Staubli VAL3: HMI_progEdit.pjx

--- HMI_progEdit.pjx ---
Parameters version=s8.12.2Cs9_BS2561 stackSize=5000 millimeterUnit=true
Program file=_bindPROG.pgx
Program file=_bindTRAJ.pgx
Program file=_btnColor.pgx
Program file=_onStartPROG.pgx
Program file=_onStartTRAJ.pgx
Program file=bind.pgx
Program file=IFedit.pgx
Program file=insertCASE.pgx
Program file=insertFOR.pgx
Program file=insertIF.pgx
Program file=insertSwitch.pgx
Program file=insetProg.pgx
Program file=main.pgx
Program file=onStart.pgx
Program file=refreshlist.pgx
Program file=resfreshPROG.pgx
Program file=resfreshTRAJ.pgx
Program file=start.pgx
Program file=stop.pgx
Program file=unbind.pgx
Data file=HMI_progEdit.dtx
Library alias=rs path=Disk://source/projectSource/robotStatus/robotStatus.pjx
Library alias=prog path=Disk://source/projectSource/program/program.pjx
Library alias=util path=Disk://HMI_cs9/HMI_util/HMI_util.pjx
Library alias=progTemp path=Disk://source/template/progTemp/progTemp.pjx
Library alias=simulate path=Disk://HMI_cs9/simulate/simulate.pjx
Library alias=trajectory path=Disk://source/projectSource/trajectory/trajectory.pjx
Library alias=io path=Disk://source/projectSource/io/io.pjx

--- HMI_progEdit.dtx ---
mdesc mNomSpeed
string sSelProg
bool bBack
public bool bBool[9]
public bool bInsert[16]
num nPageIndex
num nPageNum
public num nLstValue
string sLstValue
string sList
bool bToSave
string sPageNum
string sPageIndex
public bool bTRAJ[7]
string sPgIndexTRAJ
string sPageTRAJ
num nPgIndexTRAJ
num nPgNumTRAJ
string sTRAJList
string sInsertItem
string sPgIndexPROG
string sPagePROG
num nPgIndexPROG
num nPgNumPROG
string sPROGList
string sIFType[3]
public num nIFValue[3]
string sIFIndex[3]
string sANDOR1
string sANDOR2
bool bIFConfirm
bool bIFCancel
string sLastANDOR2
string sLastANDOR1
bool bSwitchOK
bool bSwitchCancel
string sIOList
string sSwitchValue
num nCaseValue
num nFORValue
string sForValue
bool bSelProg
bool bSelTraj
bool bBindTRAJ
bool bBindProg
num nSelType

--- main.pgx ---
public program main(string x_sSelProg)
  local bool l_bExit
  local bool l_bRefresh
  local num l_nIndex
begin
  //x_sSelProg-选中的prog
  do
    if util:sPage!="editProg"
      util:sPage="editProg"
      sSelProg= x_sSelProg
      call onStart()
      call bind()
      userPage(util:sPage)
      delay(0.5)
      l_bRefresh=true
    endIf

    if bBool[1]
      bBool[1]=false
      call simulate:simulatePROG(sSelProg)
    elseIf bBool[2]
      bBool[2]=false
      call prog:deleteProgItem(sSelProg,sLstValue,bToSave)
      l_bRefresh=true
    elseIf bBool[3]
      bBool[3]=false

    elseIf bBool[4]
      bBool[4]=false
      progTemp:libSave()
      delay(0.1)
      popUpMsg("数据已保存")
    elseIf bBool[5]
      bBool[5]=false
      nPageIndex=0
      l_bRefresh=true
    elseIf bBool[6]
      bBool[6]=false
      if nPageIndex>0
        nPageIndex=nPageIndex-1
      endIf
      l_bRefresh=true
    elseIf bBool[7]
      bBool[7]=false
      if nPageIndex<nPageNum-1
        nPageIndex=nPageIndex+1
      endIf
      l_bRefresh=true
    elseIf bBool[8]
      bBool[8]=false
      nPageIndex=nPageNum-1
      l_bRefresh=true
    elseIf bInsert[0]
      bInsert[0]=false
      call unbind()
      call prog:getProgItemIndex(sSelProg,sLstValue,l_nIndex)
      //call insetTRAJ(l_nIndex)
      l_bRefresh=true
    elseIf bInsert[1]
      bInsert[1]=false
      call unbind()
      call prog:getProgItemIndex(sSelProg,sLstValue,l_nIndex)
      call insetProg(l_nIndex,bToSave)
      l_bRefresh=true
    elseIf bInsert[2]
      bInsert[2]=false
      call insertIF()
      l_bRefresh=true
    elseIf bInsert[3]
      bInsert[3]=false
      call prog:getProgItemIndex(sSelProg,sLstValue,l_nIndex)
      call prog:insertENDIF(sSelProg,l_nIndex,bToSave)
      l_bRefresh=true
    elseIf bInsert[4]
      bInsert[4]=false
      call insertSwitch()
      l_bRefresh=true
    elseIf bInsert[5]
      bInsert[5]=false
      call prog:getProgItemIndex(sSelProg,sLstValue,l_nIndex)
      call insertCASE(l_nIndex)
      l_bRefresh=true
    elseIf bInsert[6]
      bInsert[6]=false
      call prog:getProgItemIndex(sSelProg,sLstValue,l_nIndex)
      call prog:insertENDSwitch(sSelProg,l_nIndex,bToSave)
      l_bRefresh=true
    elseIf bInsert[7]
      bInsert[7]=false
      call prog:getProgItemIndex(sSelProg,sLstValue,l_nIndex)
      call insertFOR(l_nIndex)
      l_bRefresh=true
    elseIf bBack
      bBack=false
      //call prog:onSave(bToSave)
      l_bExit=true
    endIf

    if l_bRefresh
      l_bRefresh=false
      call refreshlist()

    endIf



    delay(0)
  until l_bExit==true
  if bToSave
    call prog:onSave(bToSave)
  endIf
end

--- start.pgx ---
program start()
begin
end

--- _bindPROG.pgx ---
program _bindPROG(string x_sHtml)
  local num l_i
  local string l_sbtn
begin
  for l_i = 1 to 6
    l_sbtn="btn"+toString("",l_i)
    userPageBindClick(x_sHtml,l_sbtn,bInsert[l_i],true)
  endFor

  userPageBind(x_sHtml,"lbl1","innerHTML",sPgIndexPROG,1,"r")
  userPageBind(x_sHtml,"lbl2","innerHTML",sPagePROG,1,"r")

  userPageBindClick(x_sHtml,"btn7",bSelProg,true)
  userPageBindClick(x_sHtml,"btn8",bSelTraj,true)
  userPageBind(x_sHtml,"lst1","value",sInsertItem,1,"rw")

end

--- _bindTRAJ.pgx ---
program _bindTRAJ()
  local num l_i
  local string l_sbtn
begin
  for l_i = 1 to 6
    l_sbtn="btn"+toString("",l_i)
    userPageBindClick("insertTRAJ",l_sbtn,bInsert[l_i],true)
  endFor

  userPageBind("insertTRAJ","lbl1","innerHTML",sPgIndexTRAJ,1,"r")
  userPageBind("insertTRAJ","lbl2","innerHTML",sPageTRAJ,1,"r")


  userPageBind("insertTRAJ","lst1","value",sInsertItem,1,"rw")
end

--- _btnColor.pgx ---
public program _btnColor(num x_nSelType, string x_sHtml)
begin
  switch x_nSelType
    case 1
      userPageSet(x_sHtml,"btn7","style.backgroundColor","#7CB5FF")
      userPageSet(x_sHtml,"btn7","style.color","#FFFFFF")
      userPageSet(x_sHtml,"btn8","style.backgroundColor","#FFFFFF")
      userPageSet(x_sHtml,"btn8","style.color","#838A8F")
    break
    case 2
      userPageSet(x_sHtml,"btn8","style.backgroundColor","#7CB5FF")
      userPageSet(x_sHtml,"btn8","style.color","#FFFFFF")
      userPageSet(x_sHtml,"btn7","style.backgroundColor","#FFFFFF")
      userPageSet(x_sHtml,"btn7","style.color","#838A8F")
    break
  endSwitch

end

--- _onStartPROG.pgx ---
public program _onStartPROG(string x_sHtml)
begin
  nPgIndexPROG=0
  nPgNumPROG=0
  sPagePROG=""
  sPgIndexPROG=""
  bSelProg=true
  bSelTraj=false
  if bSelProg
    call resfreshPROG(x_sHtml)
  elseIf bSelTraj
    call resfreshTRAJ(x_sHtml)
  endIf
end

--- _onStartTRAJ.pgx ---
public program _onStartTRAJ()
begin
  nPgIndexTRAJ=0
  nPgNumTRAJ=0
  sPageTRAJ=""
  sPgIndexTRAJ=""
//  call resfreshTRAJ()
end

--- bind.pgx ---
program bind()
  local string l_sbtn
  local num l_i
begin
  //button
  userPageBindClick("editProg","btnback",bBack,true)
  for l_i = 1 to 8
    l_sbtn="btn"+toString("",l_i)
    userPageBindClick("editProg",l_sbtn,bBool[l_i],true)
  endFor

  for l_i = 0 to 8
    l_sbtn="btn1"+toString("",l_i)
    userPageBindClick("editProg",l_sbtn,bInsert[l_i],true)
  endFor

  //lbl
  userPageBind("editProg","lbl1","innerHTML",sSelProg,1,"r")
  userPageBind("editProg","lbleditindex","innerHTML",sPageIndex,1,"r")
  userPageBind("editProg","lbleditpage","innerHTML",sPageNum,1,"r")

  //lst
  userPageBind("editProg","lst1","options",sList,size(sList),"r")
  userPageBind("editProg","lst1","value",sLstValue,1,"rw")

end

--- IFedit.pgx ---
program IFedit(num x_nIndex)
begin
  call prog:editIF(sSelProg,x_nIndex,sIFType,sIFIndex,nIFValue,sANDOR1,sANDOR2,bToSave)
end

--- insertCASE.pgx ---
public program insertCASE(num x_nProgIndex)
  local bool l_bExit
  local bool l_bRefreh
  local num l_nProgIndex
  local num l_i
  local bool l_bRefresh
begin
  do
    if util:sPage!="insertCASE"
      util:sPage="insertCASE"
      call _onStartPROG(util:sPage)
      call _bindPROG(util:sPage)
      userPageBind("insertCASE","nmb1","value",nCaseValue,1,"rw")
      if size(sIOList)!=(size(io:aInItem)+1)
        resize(sIOList,1,size(io:aInItem)+1)
      endIf
      for l_i = 1 to size(sIOList)-1
        sIOList[l_i-1]=toString("",l_i-1)+","+io:aInItem[l_i-1].sComment
      endFor
      sIOList[0]=""
      userPage(util:sPage)
      delay(0.5)
    endIf

    //btn
    if bSelProg
      bSelProg=false
      nSelType=1
      l_bRefresh=true
      nPgIndexPROG=0
    elseIf bSelTraj
      bSelTraj=false
      nSelType=2
      l_bRefresh=true
      nPgIndexPROG=0
    endIf

    //refresh
    if l_bRefresh
      l_bRefresh=false
      call _btnColor(nSelType,util:sPage)
      switch nSelType
        case 1
          call resfreshPROG(util:sPage)
        break
        case 2
          nPgIndexTRAJ=0
          call resfreshTRAJ(util:sPage)
        break
      endSwitch
    endIf

    if bInsert[1]
      bInsert[1]=false

      call prog:insertCASE(sSelProg,x_nProgIndex,sInsertItem,bToSave,nCaseValue,nSelType)

      l_bExit=true
    elseIf bInsert[2]
      bInsert[2]=false
      l_bExit=true
    elseIf bInsert[3]
      bInsert[3]=false
      nPgIndexPROG=0
      l_bRefreh=true
    elseIf bInsert[4]
      bInsert[4]=false
      if nPgIndexPROG>0
        nPgIndexPROG=nPgIndexPROG-1
      endIf
      l_bRefreh=true
    elseIf bInsert[5]
      bInsert[5]=false
      if nPgIndexPROG<nPgNumPROG-1
        nPgIndexPROG=nPgIndexPROG+1
      endIf
      l_bRefreh=true
    elseIf bInsert[6]
      bInsert[6]=false
      nPgIndexPROG=nPgNumPROG-1
      l_bRefreh=true
    endIf





    delay(0)
  until l_bExit==true
end

--- insertFOR.pgx ---
public program insertFOR(num x_nProgIndex)
  local bool l_bExit
  local bool l_bRefreh
  local num l_nProgIndex
  local num l_i
  local bool l_bRefresh
begin
  do
    if util:sPage!="insertFOR"
      util:sPage="insertFOR"
      call _onStartPROG(util:sPage)
      call _bindPROG(util:sPage)
      userPageBind("insertFOR","nmb1","value",nFORValue,1,"rw")
      if size(sIOList)!=(size(io:aInItem)+1)
        resize(sIOList,1,size(io:aInItem)+1)
      endIf
      for l_i = 1 to size(sIOList)-1
        sIOList[l_i-1]=toString("",l_i-1)+","+io:aInItem[l_i-1].sComment
      endFor
      sIOList[0]="value"
      userPageBind("insertFOR","cbx1","options",sIOList,size(sIOList),"r")
      userPageBind("insertFOR","cbx1","value",sForValue,1,"rw")
      userPage(util:sPage)
      delay(0.5)
    endIf

    //btn
    if bSelProg
      bSelProg=false
      nSelType=1
      l_bRefresh=true
      nPgIndexPROG=0
    elseIf bSelTraj
      bSelTraj=false
      nSelType=2
      l_bRefresh=true
      nPgIndexPROG=0
    endIf


    //refresh
    if l_bRefresh
      l_bRefresh=false
      call _btnColor(nSelType,util:sPage)
      switch nSelType
        case 1
          call resfreshPROG(util:sPage)
        break
        case 2
          nPgIndexTRAJ=0
          call resfreshTRAJ(util:sPage)
        break
      endSwitch
    endIf

    if bInsert[1]
      bInsert[1]=false

      call prog:insertFOR(sSelProg,x_nProgIndex,sInsertItem,nFORValue,sForValue,bToSave,nSelType)

      l_bExit=true
    elseIf bInsert[2]
      bInsert[2]=false
      l_bExit=true
    elseIf bInsert[3]
      bInsert[3]=false
      nPgIndexPROG=0
      l_bRefreh=true
    elseIf bInsert[4]
      bInsert[4]=false
      if nPgIndexPROG>0
        nPgIndexPROG=nPgIndexPROG-1
        l_bRefreh=true
      endIf

    elseIf bInsert[5]
      bInsert[5]=false
      if nPgIndexPROG<nPgNumPROG-1
        nPgIndexPROG=nPgIndexPROG+1
        l_bRefreh=true
      endIf

    elseIf bInsert[6]
      bInsert[6]=false
      nPgIndexPROG=nPgNumPROG-1
      l_bRefreh=true
    endIf





    delay(0)
  until l_bExit==true
end

--- insertIF.pgx ---
program insertIF()
  local bool l_bExit
  local num l_i
  local string l_scbx
  local num l_nIndex
begin
  do
    if util:sPage!="insertIF"
      util:sPage="insertIF"
      for l_i = 0 to 2
        sIFType[l_i]=""
        sIFIndex[l_i]=""
        nIFValue[l_i]=0
        sANDOR1=""
        sANDOR2=""
        l_scbx="cbx"+toString("",l_i)
        userPageBind("insertIF",l_scbx,"value",sIFType[l_i],1,"rw")
        l_scbx="cbx1"+toString("",l_i)
        userPageBind("insertIF",l_scbx,"value",sIFIndex[l_i],1,"rw")
        l_scbx="nmb"+toString("",l_i)
        userPageBind("insertIF",l_scbx,"value",nIFValue[l_i],1,"rw")

        userPageBind("insertIF","cbx7","value",sANDOR1,1,"rw")
        userPageBind("insertIF","cbx8","value",sANDOR2,1,"rw")
        userPageBindClick("insertIF","btn1",bIFConfirm,true)
        userPageBindClick("insertIF","btn2",bIFCancel,true)

      endFor
      sLastANDOR1=""
      sLastANDOR2=""
      //      userPageSet("insertIF","cbx1","disabled",true)
      //      userPageSet("insertIF","cbx2","disabled",true)
      //      userPageSet("insertIF","cbx11","disabled",true)
      //      userPageSet("insertIF","cbx12","disabled",true)
      //      userPageSet("insertIF","nmb1","disabled",true)
      //      userPageSet("insertIF","nmb1","disabled",true)
      userPage(util:sPage)
      delay(0.5)
    endIf

    //    if sLastANDOR1!=sANDOR1
    //      sLastANDOR1=sANDOR1
    //      if sANDOR1=""
    //        userPageSet("insertIF","cbx1","disabled",true)
    //        userPageSet("insertIF","cbx11","disabled",true)
    //        userPageSet("insertIF","nmb1","disabled",true)
    //        userPageSet("insertIF","cbx8","disabled",true)
    //      endIf
    //    endIf


    //button
    if bIFConfirm
      bIFConfirm=false
      call prog:getProgItemIndex(sSelProg,sLstValue,l_nIndex)
      call IFedit(l_nIndex)
      l_bExit=true
    elseIf bIFCancel
      bIFCancel=false
      l_bExit=true
    endIf



  until l_bExit==true

end

--- insertSwitch.pgx ---
program insertSwitch()
  local bool l_bExit
  local num l_i
  local num l_nIndex
  local num l_nValue
  local bool l_bResult
begin
  do
    if util:sPage!="insertSwitch"
      util:sPage="insertSwitch"
      if size(sIOList)!=(size(io:aInItem)+1)
        resize(sIOList,1,size(io:aInItem)+1)
      endIf

      for l_i = 1 to size(sIOList)-1
        sIOList[l_i-1]=toString("",l_i-1)+","+io:aInItem[l_i-1].sComment
      endFor

      sIOList[0]=""
      userPageBind("insertSwitch","cbx1","options",sIOList,size(sIOList),"r")
      userPageBind("insertSwitch","cbx1","value",sSwitchValue,1,"rw")
      userPageBindClick("insertSwitch","btn1",bSwitchOK,true)
      userPageBindClick("insertSwitch","btn2",bSwitchCancel,true)
      userPage(util:sPage)
      delay(0.5)
    endIf
    //cbx

    //button
    if bSwitchOK
      bSwitchOK=false
      call prog:getProgItemIndex(sSelProg,sLstValue,l_nIndex)
      if sSwitchValue!=""
        call prog:insertSwitch(sSelProg,l_nIndex,sSwitchValue,bToSave)
      else
        userPageAlert("请选择正确的switch值")
      endIf
      l_bExit=true
    elseIf bSwitchCancel
      bSwitchCancel=false
      l_bExit=true
    endIf




  until l_bExit==true
  l_bExit=false
end

--- insetProg.pgx ---
public program insetProg(num x_nProgIndex, bool& x_bToSave)
  local bool l_bExit
  local bool l_bRefresh
  local num l_nProgIndex
  local num l_num
  local bool l_bResult
begin
  do
    if util:sPage!="insertPROG"
      util:sPage="insertPROG"
      call _onStartPROG(util:sPage)
      call _bindPROG(util:sPage)
      userPage(util:sPage)
      delay(0.5)
    endIf

    //btn
    if bSelProg
      bSelProg=false
      nSelType=1
      l_bRefresh=true
      nPgIndexPROG=0
    elseIf bSelTraj
      bSelTraj=false
      nSelType=2
      l_bRefresh=true
      nPgIndexPROG=0
    endIf

    //refresh
    if l_bRefresh
      l_bRefresh=false
      call _btnColor(nSelType,util:sPage)
      switch nSelType
        case 1
          call resfreshPROG(util:sPage)
        break
        case 2
          nPgIndexTRAJ=0
          call resfreshTRAJ(util:sPage)
        break
      endSwitch
    endIf
    //insert btn
    if bInsert
      bInsert=false

    elseIf bInsert[1]
      bInsert[1]=false
      if nSelType==1
        call prog:insertPROG(sSelProg,x_nProgIndex,sInsertItem,x_bToSave)
      elseIf nSelType==2
        call prog:insertTRAJ(sSelProg,x_nProgIndex,sInsertItem,x_bToSave)
      endIf
      l_bExit=true
    elseIf bInsert[2]
      bInsert[2]=false
      l_bExit=true
    elseIf bInsert[3]
      bInsert[3]=false
      nPgIndexPROG=0
      l_bRefresh=true
    elseIf bInsert[4]
      bInsert[4]=false
      if nPgIndexPROG>0
        nPgIndexPROG=nPgIndexPROG-1
      endIf
      l_bRefresh=true
    elseIf bInsert[5]
      bInsert[5]=false
      if nPgIndexPROG<nPgNumPROG-1
        nPgIndexPROG=nPgIndexPROG+1
      endIf
      l_bRefresh=true
    elseIf bInsert[6]
      bInsert[6]=false
      nPgIndexPROG=nPgNumPROG-1
      l_bRefresh=true
    endIf


    delay(0)
  until l_bExit==true

end

--- onStart.pgx ---
public program onStart()
  local num l_nSize
  local string l_sMsg
  local num l_i
begin
  sLstValue=""
  nPageIndex=0
  nPageNum=1
  call refreshlist()

  sPageIndex=toString("",nPageIndex+1)
  sPageNum=toString("",nPageNum)
end

--- refreshlist.pgx ---
public program refreshlist()
  local num l_nSize
  local num l_i
  local num l_nSize1
  local string l_sMsg
  local num l_nIndex
begin
  //bulid list
  call prog:getProgItemSize(sSelProg,l_nSize)
  resize(sList,1,l_nSize)
  //npage
  if l_nSize<50
    nPageNum=1
  else
    nPageNum=roundUp(l_nSize/49)
  endIf
  //pageindex
  if nPageIndex>nPageNum-1
    nPageIndex=nPageNum-1
  endIf
  //
  if nPageIndex==(nPageNum-1)
    l_nSize1=l_nSize%49
    if l_nSize1==0
      resize(sList,1,49)
      for l_i = 0 to size(sList)-1
        call prog:pointToString(l_sMsg,sSelProg,l_i)
        sList[l_i]=toString("",l_i)+l_sMsg
      endFor
    else
      resize(sList,1,l_nSize1)
      for l_i = 0 to l_nSize1-1
        l_nIndex=nPageIndex*49+l_i
        call prog:pointToString(l_sMsg,sSelProg,l_nIndex)
        sList[l_i]=toString("",l_nIndex)+l_sMsg
      endFor
    endIf
  else
    resize(sList,1,49)
    for l_i = 0 to size(sList)-1
      call prog:pointToString(l_sMsg,sSelProg,l_i)
      sList[l_i]=toString("",l_i)+l_sMsg
    endFor
  endIf
  userPageBind("editProg","lst1","options",sList,size(sList),"r")
  sPageIndex=toString("",nPageIndex+1)
  sPageNum=toString("",nPageNum)
end

--- resfreshPROG.pgx ---
program resfreshPROG(string x_sHtml)
  local num l_nSize
  local num l_nSize1
  local num l_i
begin
  //call PROGectory:getSize(l_nSize)
  //  call PROGectory:getPROGList(sPROGList)
  call prog:getSize(l_nSize)
  call prog:getProgList(sPROGList)

  if l_nSize>49
    nPgNumPROG=roundUp(l_nSize/49)
  else
    nPgNumPROG=1
  endIf

  l_nSize1=l_nSize%49

  if nPgIndexPROG==nPgNumPROG-1
    if l_nSize1!=0
      resize(sList,1,l_nSize1)
      for l_i = 0 to size(sList)-1
        sList[l_i]=sPROGList[l_i+nPgIndexPROG*49]
      endFor
    else
      resize(sList,1,49)
      for l_i = 0 to size(sList)-1
        sList[l_i]=sPROGList[l_i+nPgIndexPROG*49]
      endFor
    endIf
  else
    resize(sList,1,49)
    for l_i = 0 to size(sList)-1
      sList[l_i]=sPROGList[l_i+nPgIndexPROG*49]
    endFor
  endIf
  userPageBind(x_sHtml,"lst1","options",sList,size(sList),"r")
  sPagePROG=toString("",nPgNumPROG)
  sPgIndexPROG=toString("",nPgIndexPROG+1)
end

--- resfreshTRAJ.pgx ---
program resfreshTRAJ(string x_sHtml)
  local num l_nSize
  local num l_nSize1
  local num l_i
begin
  call trajectory:getSize(l_nSize)
  call trajectory:getTrajList(sTRAJList)

  if l_nSize>49
    nPgNumPROG=roundUp(l_nSize/49)
  else
    nPgNumPROG=1
  endIf

  l_nSize1=l_nSize%49

  if nPgIndexPROG==nPgNumPROG-1
    if l_nSize1!=0
      resize(sList,1,l_nSize1)
      for l_i = 0 to size(sList)-1
        sList[l_i]=sTRAJList[l_i+nPgIndexPROG*49]
      endFor
    else
      resize(sList,1,49)
      for l_i = 0 to size(sList)-1
        sList[l_i]=sTRAJList[l_i+nPgIndexPROG*49]
      endFor
    endIf
  else
    resize(sList,1,49)
    for l_i = 0 to size(sList)-1
      sList[l_i]=sTRAJList[l_i+nPgIndexPROG*49]
    endFor
  endIf
  userPageBind(x_sHtml,"lst1","options",sList,size(sList),"r")
  sPagePROG=toString("",nPgNumPROG)
  sPgIndexPROG=toString("",nPgIndexPROG+1)
end

--- stop.pgx ---
program stop()
begin
end

--- unbind.pgx ---
program unbind()
begin
  userPageUnbind("editProg","lst1","value")
  userPageUnbind("editProg","lst1","options")
end
